(* IEC 61131-3 sources: ZPLC/conformance/lng, 23 files *)

(* ---- lng-008-fbd-calls-a-user-function-scale.st ---- *)
FUNCTION Scale : INT
VAR_INPUT Value : INT; Gain : INT; END_VAR
  Scale := Value * Gain;
END_FUNCTION

(* ---- lng-008-fbd-calls-a-user-function-block-latch.st ---- *)
FUNCTION_BLOCK Latch
VAR_INPUT Set : BOOL; END_VAR
VAR_OUTPUT Q : BOOL; END_VAR
  IF Set THEN
    Q := TRUE;
  END_IF;
END_FUNCTION_BLOCK

(* ---- lng-008-ld-places-a-user-function-block-hold.st ---- *)
FUNCTION_BLOCK Hold
VAR_INPUT Trigger : BOOL; END_VAR
VAR_OUTPUT Active : BOOL; END_VAR
  IF Trigger THEN
    Active := TRUE;
  END_IF;
END_FUNCTION_BLOCK

(* ---- lng-003-il-compiler-error-names-the-il-line.il ---- *)
PROGRAM Wrong
VAR
  T : TON;
  Lamp AT %QX0.0 : BOOL;
END_VAR
  LD TRUE
  CAL T(IN := 5)
  LD T.Q
  ST Lamp
END_PROGRAM

(* ---- lng-017-il-unbalanced-closing-parenthesis.il ---- *)
PROGRAM Closing
VAR
  A : BOOL;
  B : BOOL;
  X : BOOL;
END_VAR
  LD A
  AND( B
  )
  )
  ST X
END_PROGRAM

(* ---- lng-017-il-unknown-mnemonic.il ---- *)
PROGRAM Typo
VAR
  A : BOOL;
  X : BOOL;
END_VAR
  LD A
  ANDD A
  ST X
END_PROGRAM

(* ---- lng-018-il-backward-jump-loop.il ---- *)
PROGRAM Loop
VAR
  I : INT;
  Out AT %QW0 : INT;
END_VAR
  LD 0
  ST I
again:
  LD I
  ADD 1
  ST I
  LT 3
  JMPC again
  LD I
  ST Out
END_PROGRAM

(* ---- lng-018-il-conditional-jump-follows-input.il ---- *)
PROGRAM Skip
VAR
  Go AT %IX0.0 : BOOL;
  Ran AT %QW0 : INT;
  Passed AT %QW1 : INT;
END_VAR
  LD Go
  JMPCN done
  LD Ran
  ADD 1
  ST Ran
done:
  LD Passed
  ADD 1
  ST Passed
END_PROGRAM

(* ---- lng-018-il-duplicate-label.il ---- *)
PROGRAM TwoLabels
VAR
  A : BOOL;
  X : BOOL;
END_VAR
again:
  LD A
  ST X
again:
  LD X
  ST A
END_PROGRAM

(* ---- lng-018-il-jump-runs-every-scan.il ---- *)
PROGRAM JumpTest
VAR
  A : BOOL;
  Hits AT %QW0 : INT;
  Tail AT %QW1 : INT;
END_VAR
  LD Hits
  ADD 1
  ST Hits
  LD A
  JMPC skip
  LD Tail
  ADD 1
  ST Tail
skip:
  LD Hits
  ST Hits
END_PROGRAM

(* ---- lng-018-il-jump-to-unknown-label.il ---- *)
PROGRAM BadLabel
VAR
  A : BOOL;
  X : BOOL;
END_VAR
  LD A
  JMPC nowhere
  ST X
END_PROGRAM

(* ---- lng-018-il-unconditional-jump-to-unknown-label.il ---- *)
PROGRAM BadJump
VAR
  X : BOOL;
END_VAR
  LD TRUE
  ST X
  JMP missing
END_PROGRAM

(* ---- lng-019-il-arithmetic-in-parentheses.il ---- *)
PROGRAM Scaled
VAR
  Out AT %QW0 : INT;
  Cmp AT %QX2.0 : BOOL;
END_VAR
  LD 10
  MUL( 2
  ADD 3
  )
  ST Out
  GT( 40
  ADD 5
  )
  ST Cmp
END_PROGRAM

(* ---- lng-019-il-conditional-call-and-return.il ---- *)
PROGRAM Calls
VAR
  Call AT %IX0.0 : BOOL;
  Skip AT %IX0.1 : BOOL;
  OnTrue : RS;
  OnFalse : RS;
  Ran AT %QW1 : INT;
  A AT %QX0.0 : BOOL;
  B AT %QX0.1 : BOOL;
END_VAR
  LD Call
  CALC OnTrue(S := TRUE, R1 := FALSE)
  LD Skip
  CALCN OnFalse(S := TRUE, R1 := FALSE)
  LD OnTrue.Q1
  ST A
  LD OnFalse.Q1
  ST B
  LD Call
  RETC
  LD Ran
  ADD 1
  ST Ran
END_PROGRAM

(* ---- lng-019-il-direct-address-operands.il ---- *)
PROGRAM Direct
  LD %IX0.0
  ANDN %IX0.1
  ST %QX0.0
END_PROGRAM

(* ---- lng-019-il-negated-operators-set-and-reset.il ---- *)
PROGRAM Negated
VAR
  A AT %IX0.0 : BOOL;
  B AT %IX0.1 : BOOL;
  X AT %QX0.0 : BOOL;
  Y AT %QX0.1 : BOOL;
  Latch AT %QX0.2 : BOOL;
END_VAR
  LDN A
  ANDN B
  ST X
  STN Y
  LD A
  S Latch
  LD B
  R Latch
END_PROGRAM

(* ---- lng-019-il-nested-parentheses.il ---- *)
PROGRAM Nested
VAR
  A AT %IX0.0 : BOOL;
  B AT %IX0.1 : BOOL;
  C AT %IX0.2 : BOOL;
  D AT %IX0.3 : BOOL;
  X AT %QX0.0 : BOOL;
END_VAR
  LD A
  OR( B
  AND( C
  ORN D )
  )
  ST X
END_PROGRAM

(* ---- lng-019-il-parenthesised-operation.il ---- *)
PROGRAM Parens
VAR
  A : BOOL;
  B : BOOL;
  C : BOOL := TRUE;
  X AT %QX0.0 : BOOL;
END_VAR
  LD A
  AND( B
  OR C
  )
  ST X
END_PROGRAM

(* ---- lng-019-il-real-accumulator.il ---- *)
PROGRAM RealSum
VAR
  R1 : REAL := 1.5;
  R2 AT %QD0 : REAL;
END_VAR
  LD R1
  ADD 2.25
  ST R2
END_PROGRAM

(* ---- lng-019-il-real-arithmetic-and-comparison.il ---- *)
PROGRAM RealMath
VAR
  A : REAL := 6.0;
  Big AT %QX4.0 : BOOL;
  Quot AT %QD0 : REAL;
END_VAR
  LD A
  DIV 4.0
  MUL 3
  SUB 0.5
  ST Quot
  GT 3.5
  ST Big
END_PROGRAM

(* ---- lng-019-il-time-accumulator.il ---- *)
PROGRAM Times
VAR
  Total AT %QD0 : TIME;
END_VAR
  LD T#1s
  ADD T#500ms
  ST Total
END_PROGRAM

(* ---- lng-020-il-load-and-store.il ---- *)
PROGRAM Gate
VAR
  A AT %IX0.0 : BOOL;
  B AT %IX0.1 : BOOL;
  X AT %QX0.0 : BOOL;
END_VAR
  LD A
  AND B
  ST X
END_PROGRAM

(* ---- lng-020-il-remaining-operators.il ---- *)
PROGRAM Rest
VAR
  A AT %IX0.0 : BOOL;
  B AT %IX0.1 : BOOL;
  Xor1 AT %QX0.0 : BOOL;
  Xor2 AT %QX0.1 : BOOL;
  Not1 AT %QX0.2 : BOOL;
  IsEq AT %QX0.3 : BOOL;
  IsNe AT %QX0.4 : BOOL;
  IsGe AT %QX0.5 : BOOL;
  IsLe AT %QX0.6 : BOOL;
  Remainder AT %QW1 : INT;
  Negated AT %QW2 : INT;
  Rises AT %QW3 : INT;
  Hit AT %QW4 : INT;
  N : INT := 7;
  Cnt : CTU;
END_VAR
  LD A
  XOR B
  ST Xor1
  LD A
  XORN B
  ST Xor2
  LD A
  NOT
  ST Not1
  LD N
  EQ 7
  ST IsEq
  LD N
  NE 7
  ST IsNe
  LD N
  GE 8
  ST IsGe
  LD N
  LE 7
  ST IsLe
  LD N
  MOD 4
  ST Remainder
  LD N
  NEG
  ST Negated
  CAL Cnt(CU := A, R := FALSE, PV := 100)
  LD Cnt.CV
  ST Rises
  JMP skip
  LD 99
  ST Hit
skip:
  LD 1
  ST Hit
  RET
  LD 77
  ST Hit
END_PROGRAM
